Yaskawa INFORM job: MOVEUNTI.JBI

/JOB
//NAME MOVEUNTI
//POS
///NPOS 0,0,0,2,0,0
///TOOL 0
///POSTYPE BASE
///RECTAN
///RCONF 1,0,0,0,1,0,0,0
P0002=1529.187,-331.251,500.000,180.00,0.00,90.00
///RCONF 0,0,0,0,0,0,0,0
P0003=0.000,0.000,-600.000,0.00,0.00,0.00
//INST
///DATE 2026/10/27 16:26
///ATTR SC,RW
///GROUP1 RB1
NOP
MOVL P002 V=I000 PL=0 DEC=50
IMOV P003 V=120.0 PL=0 BF UNTIL IN#(1)=ON
HAND HNO: 2 ON
END
